(* IEC 61131-3 sources: llm-plc-st-eval/codesys/dobles/A4, 8 files *)

(* ---- 01_Correcta.st ---- *)
(* DOBLE DE PRUEBA A4/Correcta - NO ES CORPUS. Esperado: veredicto 1 *)
FUNCTION_BLOCK FB_Rampa
VAR_INPUT
    SPvel : REAL;
    paroRapido : BOOL;
    ciclo : TIME;
END_VAR
VAR_OUTPUT
    CVvel : REAL;
END_VAR
VAR
    d : REAL;
    obj : REAL;
    bajada : REAL;
    llego : BOOL;
END_VAR
d := TIME_TO_REAL(ciclo) / 1000.0;
IF paroRapido THEN
    obj := 0.0;
    bajada := 40.0;
ELSE
    obj := SPvel;
    bajada := 20.0;
END_IF
IF CVvel < obj THEN
    CVvel := MIN(obj, CVvel + 10.0 * d);
ELSIF CVvel > obj THEN
    CVvel := MAX(obj, CVvel - bajada * d);
END_IF
END_FUNCTION_BLOCK

(* ---- 02_SubidaRapida.st ---- *)
(* DOBLE DE PRUEBA A4/SubidaRapida - NO ES CORPUS. Esperado: veredicto 2, falla en el paso 2 *)
FUNCTION_BLOCK FB_Rampa
VAR_INPUT
    SPvel : REAL;
    paroRapido : BOOL;
    ciclo : TIME;
END_VAR
VAR_OUTPUT
    CVvel : REAL;
END_VAR
VAR
    d : REAL;
    obj : REAL;
    bajada : REAL;
    llego : BOOL;
END_VAR
d := TIME_TO_REAL(ciclo) / 1000.0;
IF paroRapido THEN
    obj := 0.0;
    bajada := 40.0;
ELSE
    obj := SPvel;
    bajada := 20.0;
END_IF
IF CVvel < obj THEN
    CVvel := MIN(obj, CVvel + 20.0 * d);
ELSIF CVvel > obj THEN
    CVvel := MAX(obj, CVvel - bajada * d);
END_IF
END_FUNCTION_BLOCK

(* ---- 03_BajadaLenta.st ---- *)
(* DOBLE DE PRUEBA A4/BajadaLenta - NO ES CORPUS. Esperado: veredicto 2, falla en el paso 4 *)
FUNCTION_BLOCK FB_Rampa
VAR_INPUT
    SPvel : REAL;
    paroRapido : BOOL;
    ciclo : TIME;
END_VAR
VAR_OUTPUT
    CVvel : REAL;
END_VAR
VAR
    d : REAL;
    obj : REAL;
    bajada : REAL;
    llego : BOOL;
END_VAR
d := TIME_TO_REAL(ciclo) / 1000.0;
IF paroRapido THEN
    obj := 0.0;
    bajada := 40.0;
ELSE
    obj := SPvel;
    bajada := 10.0;
END_IF
IF CVvel < obj THEN
    CVvel := MIN(obj, CVvel + 10.0 * d);
ELSIF CVvel > obj THEN
    CVvel := MAX(obj, CVvel - bajada * d);
END_IF
END_FUNCTION_BLOCK

(* ---- 04_ParoLento.st ---- *)
(* DOBLE DE PRUEBA A4/ParoLento - NO ES CORPUS. Esperado: veredicto 2, falla en el paso 7 *)
FUNCTION_BLOCK FB_Rampa
VAR_INPUT
    SPvel : REAL;
    paroRapido : BOOL;
    ciclo : TIME;
END_VAR
VAR_OUTPUT
    CVvel : REAL;
END_VAR
VAR
    d : REAL;
    obj : REAL;
    bajada : REAL;
    llego : BOOL;
END_VAR
d := TIME_TO_REAL(ciclo) / 1000.0;
IF paroRapido THEN
    obj := 0.0;
    bajada := 20.0;
ELSE
    obj := SPvel;
    bajada := 20.0;
END_IF
IF CVvel < obj THEN
    CVvel := MIN(obj, CVvel + 10.0 * d);
ELSIF CVvel > obj THEN
    CVvel := MAX(obj, CVvel - bajada * d);
END_IF
END_FUNCTION_BLOCK

(* ---- 05_ParoInstantaneo.st ---- *)
(* DOBLE DE PRUEBA A4/ParoInstantaneo - NO ES CORPUS. Esperado: veredicto 2, falla en el paso 7 *)
FUNCTION_BLOCK FB_Rampa
VAR_INPUT
    SPvel : REAL;
    paroRapido : BOOL;
    ciclo : TIME;
END_VAR
VAR_OUTPUT
    CVvel : REAL;
END_VAR
VAR
    d : REAL;
    obj : REAL;
    bajada : REAL;
    llego : BOOL;
END_VAR
d := TIME_TO_REAL(ciclo) / 1000.0;
IF paroRapido THEN
    obj := 0.0;
    bajada := 40.0;
ELSE
    obj := SPvel;
    bajada := 20.0;
END_IF
IF paroRapido THEN
    CVvel := 0.0;
END_IF
IF CVvel < obj THEN
    CVvel := MIN(obj, CVvel + 10.0 * d);
ELSIF CVvel > obj THEN
    CVvel := MAX(obj, CVvel - bajada * d);
END_IF
END_FUNCTION_BLOCK

(* ---- 06_ParoNoMantiene.st ---- *)
(* DOBLE DE PRUEBA A4/ParoNoMantiene - NO ES CORPUS. Esperado: veredicto 2, falla en el paso 8 *)
FUNCTION_BLOCK FB_Rampa
VAR_INPUT
    SPvel : REAL;
    paroRapido : BOOL;
    ciclo : TIME;
END_VAR
VAR_OUTPUT
    CVvel : REAL;
END_VAR
VAR
    d : REAL;
    obj : REAL;
    bajada : REAL;
    llego : BOOL;
END_VAR
d := TIME_TO_REAL(ciclo) / 1000.0;
IF paroRapido THEN
    obj := 0.0;
    bajada := 40.0;
ELSE
    obj := SPvel;
    bajada := 20.0;
END_IF
IF NOT paroRapido THEN
    llego := FALSE;
END_IF
IF paroRapido AND llego THEN
    obj := SPvel;
    bajada := 20.0;
END_IF
IF CVvel < obj THEN
    CVvel := MIN(obj, CVvel + 10.0 * d);
ELSIF CVvel > obj THEN
    CVvel := MAX(obj, CVvel - bajada * d);
END_IF
IF paroRapido AND CVvel <= 0.0 THEN
    llego := TRUE;
END_IF
END_FUNCTION_BLOCK

(* ---- 07_Sobrepaso.st ---- *)
(* DOBLE DE PRUEBA A4/Sobrepaso - NO ES CORPUS. Esperado: veredicto 2, falla en el paso 0 *)
FUNCTION_BLOCK FB_Rampa
VAR_INPUT
    SPvel : REAL;
    paroRapido : BOOL;
    ciclo : TIME;
END_VAR
VAR_OUTPUT
    CVvel : REAL;
END_VAR
VAR
    d : REAL;
    obj : REAL;
    bajada : REAL;
    llego : BOOL;
END_VAR
d := TIME_TO_REAL(ciclo) / 1000.0;
IF paroRapido THEN
    obj := 0.0;
    bajada := 40.0;
ELSE
    obj := SPvel;
    bajada := 20.0;
END_IF
IF CVvel < obj THEN
    CVvel := CVvel + 10.0 * d;
ELSIF CVvel > obj THEN
    CVvel := CVvel - bajada * d;
END_IF
END_FUNCTION_BLOCK

(* ---- 08_CicloEnMs.st ---- *)
(* DOBLE DE PRUEBA A4/CicloEnMs - NO ES CORPUS. Esperado: veredicto 2, falla en el paso 2 *)
FUNCTION_BLOCK FB_Rampa
VAR_INPUT
    SPvel : REAL;
    paroRapido : BOOL;
    ciclo : TIME;
END_VAR
VAR_OUTPUT
    CVvel : REAL;
END_VAR
VAR
    d : REAL;
    obj : REAL;
    bajada : REAL;
    llego : BOOL;
END_VAR
d := TIME_TO_REAL(ciclo);
IF paroRapido THEN
    obj := 0.0;
    bajada := 40.0;
ELSE
    obj := SPvel;
    bajada := 20.0;
END_IF
IF CVvel < obj THEN
    CVvel := MIN(obj, CVvel + 10.0 * d);
ELSIF CVvel > obj THEN
    CVvel := MAX(obj, CVvel - bajada * d);
END_IF
END_FUNCTION_BLOCK
